// TwinCAT 3 PLC project PannenkoekSysteem
// ProgramVersion: 3.1.4026.20
// CompilerDefines: VISU_USEPROPERTYINFO
// libraries:
//   Tc2_Standard, * (Beckhoff Automation GmbH)
//   Tc2_System, * (Beckhoff Automation GmbH)
//   Tc3_IotBase, * (Beckhoff Automation GmbH)
//   Tc3_Module, * (Beckhoff Automation GmbH)
//   Tc3_Vision, * (Beckhoff Automation GmbH)
// project tree:
//   DUTs/ E_MainState.TcDUT
//   / GlobalTextList.TcGTLO, PlcTask.TcTTO, Visualization Manager.TcVMO (not stored)
//   GVLs/ GVL_Config.TcGVL, GVL_Data.TcGVL, GVL_Inputs.TcGVL, GVL_MQTT.TcGVL, GVL_Outputs.TcGVL
//   POUs/ FB_MQTT.TcPOU, FB_QrVision.TcPOU, F_ParseErrorDisplay.TcPOU, F_ParseStateDisplay.TcPOU, FB_StateMachine.TcPOU, FB_Transportband.TcPOU, MAIN.TcPOU
//   VISUs/ PannenkoekenDashboard.TcVIS
// real-time tasks:
//   TASK PlcTask: cycle T#10ms, priority 20, ADS port 350
//   TASK VnTask ImgAcq (Camera1): cycle T#1ms, priority 5, ADS port 351
//   TASK VnTask ADS (Camera1): cycle T#10ms, priority 6, ADS port 352
// motion (NC):
//   TASK NC-Task 1 SAF: cycle T#2ms, priority 4, ADS port 501
//   TASK NC-Task 1 SVB: cycle T#10ms, priority 8, ADS port 511
//   AXIS Axis 1 (id 1)
//     Dynamic: AccelerationMaximum=200, DecelerationMaximum=200
//     Velo: SlowManual=5, FastManual=20, Maximum=50
//     MotionControl: Range=500, Time=20
//     OtherSettings: AllowMotionCmdToSlave=true
//     encoder EncType=4
//       EncPara: EncMode=1, MaxCount=#x0000ffff
//     drive DrvType=23
//       Analog: VeloReferenz=50, TorqueSetpointScale=10, ScaleFactorActTorque=0.1
//       TimeComp: TaskDelayCycles=1
//     controller CtrType=1
//       CtrPara: PriorControlFactor=1
//         PosDiffControl: Range=20000
//         Observer: BandWidth=20
// I/O:
//   DEVICE Device 2 (EtherCAT), AmsNetId 172.18.237.156.3.1
//     Term 1 (EK1100) [EK1100 EtherCAT Coupler (2A E-Bus)]
//       Term 2 (EL7332) [EL7332 2Ch. DC motor output stage (24V, 1.5A)]
//       Term 3 (EL6001) [EL6001 Interface (RS232)]
//       Box 4 (BK1250)
//   DEVICE Device 1 (RT-Ethernet Adapter)
// variable links:
//   NC-Task 1 SAF/Axes/Axis 1 <-> Device 2 (EtherCAT)/Term 1 (EK1100)/Term 2 (EL7332)
//     Drive/Inputs/In/nState1 @bit 3 <-> DCM Status Channel 1/Status/Error
//     Drive/Inputs/In/nState1 @bit 5 <-> DCM Status Channel 1/Status/Moving negative
//     Drive/Inputs/In/nState1 @bit 4 <-> DCM Status Channel 1/Status/Moving positive
//     Drive/Inputs/In/nState1 @bit 1 <-> DCM Status Channel 1/Status/Ready
//     Drive/Inputs/In/nState1 <-> DCM Status Channel 1/Status/Ready to enable
//     Drive/Inputs/In/nState1 @bit 6 <-> DCM Status Channel 1/Status/Torque reduced
//     Drive/Inputs/In/nState1 @bit 2 <-> DCM Status Channel 1/Status/Warning
//     Drive/Inputs/In/nState2 @bit 3 <-> DCM Status Channel 1/Status/Digital input 1
//     Drive/Inputs/In/nState2 @bit 4 <-> DCM Status Channel 1/Status/Digital input 2
//     Drive/Inputs/In/nState2 @bit 5 <-> DCM Status Channel 1/Status/Sync error
//     Drive/Inputs/In/nState2 @bit 7 <-> DCM Status Channel 1/Status/TxPDO Toggle
//     Drive/Inputs/In/nState4 @bit 1 <-> WcState/InputToggle
//     Drive/Inputs/In/nState4 <-> WcState/WcState
//     Drive/Outputs/Out/nCtrl1 <-> DCM Control Channel 1/Control/Enable
//     Drive/Outputs/Out/nCtrl1 @bit 2 <-> DCM Control Channel 1/Control/Reduce torque
//     Drive/Outputs/Out/nCtrl1 @bit 1 <-> DCM Control Channel 1/Control/Reset
//     Drive/Outputs/Out/nDataOut2[0] <-> DCM Velocity Channel 1/Velocity

CONFIGURATION PannenkoekSysteem
    RESOURCE PLC ON TwinCAT3
        TASK PlcTask(INTERVAL := T#10ms, PRIORITY := 20);
        PROGRAM MAIN WITH PlcTask : MAIN;
    END_RESOURCE
END_CONFIGURATION

// ---- DUTs/E_MainState.TcDUT
{attribute 'qualified_only'}
{attribute 'strict'}
TYPE E_MainState :
(
    INIT,
    IDLE,
    ERROR,
    SEQ_WAIT_START,
    SEQ_FEED_BLOCK,
    SEQ_MOVE_CAMERA,
    SEQ_WAIT_CAMERA,
    SEQ_SCAN_CAMERA,
    SEQ_MOVE_SCALE,
    SEQ_WAIT_SCALE,
    SEQ_MOVE_MIXER,
    SEQ_WAIT_MIXER,
    SEQ_MOVE_INDUCTIVE,
    SEQ_WAIT_INDUCTIVE,
    SEQ_MOVE_DISCARD,
    SEQ_WAIT_DISCARD,
    SEQ_COMPLETE,
    SEQ_ERROR
);
END_TYPE

// ---- GVLs/GVL_Config.TcGVL
{attribute 'qualified_only'}
VAR_GLOBAL
  bAutoSequenceEnable : BOOL := TRUE;      // Master switch for the automated line sequence
  tFeedDuration       : TIME := T#3S;      // Conveyor run time before the robot starts
  tRobotTimeout       : TIME := T#20S;     // Max time to wait for a robot move
  tQrScanDuration     : TIME := T#5S;      // Max time to scan the block at the camera
  tSensorWaitDuration : TIME := T#5S;      // Max time to wait for the inductive sensor

  sPoseCamera    : STRING(32) := 'camera';
  sPoseScale     : STRING(32) := 'scale';
  sPoseMixer     : STRING(32) := 'mixer';
  sPoseInductive : STRING(32) := 'inductive';
  sPoseDiscard   : STRING(32) := 'discard';
END_VAR

// ---- GVLs/GVL_Data.TcGVL
{attribute 'qualified_only'}
VAR_GLOBAL
  bQrEnabled     : BOOL := FALSE;
  bQrCodeFound   : BOOL := FALSE;
  bQrCameraConnected : BOOL := FALSE; // Camera hardware connected
  bQrActive      : BOOL := FALSE;    // Enabled OR camera connected (VISU lamp)
  sQrCodeText    : STRING(255) := '';
  sQrDisplayText : STRING(512) := 'QR scanner OFF';
  hrQrVision     : HRESULT := 0;
END_VAR

// ---- GVLs/GVL_Inputs.TcGVL
{attribute 'qualified_only'}
  VAR_GLOBAL
  END_VAR

// ---- GVLs/GVL_MQTT.TcGVL
{attribute 'qualified_only'}
VAR_GLOBAL
	// MQTT Broker Configuration - HiveMQ Public Broker
	sMqttBroker			: STRING(255) := '192.168.0.198';	// MQTT broker address
	nMqttPort			: UINT := 1883;						// Standard MQTT port
	sMqttClientID		: STRING(255) := 'Twincat_Test'; // Unique client ID
	bEnableMqtt			: BOOL := TRUE;						// Enable/disable MQTT connection
	
	// MQTT Topics - Robot
	sTopicRobotCmd			: STRING(255) := 'pancake/robot/cmd';
	sTopicRobotState		: STRING(255) := 'pancake/robot/state';
	sTopicRobotError		: STRING(255) := 'pancake/robot/error';
	sTopicRobotHeartbeat	: STRING(255) := 'pancake/robot/heartbeat';

	// MQTT Topics - Transportband
	sTopicTransportbandCmd		: STRING(255) := 'pancake/transportband/cmd';
	sTopicTransportbandState	: STRING(255) := 'pancake/transportband/state';
	sTopicTransportbandError	: STRING(255) := 'pancake/transportband/error';

	// MQTT Topics - Mixer
	sTopicMixerCmd				: STRING(255) := 'pancake/mixer/cmd';
	sTopicMixerState			: STRING(255) := 'pancake/mixer/state';
	sTopicMixerError			: STRING(255) := 'pancake/mixer/error';
	
	bVisuStartTransportband : BOOL := FALSE;				// VISU button - Start transportband
	bVisuStopTransportband	: BOOL := FALSE;				// VISU button - Stop transportband
	bVisuStartSequence		: BOOL := FALSE;				// VISU button - Start automated sequence
	bVisuAutoSequenceEnable	: BOOL := TRUE;				// VISU toggle - Automatic line sequence
	
	bVisuStartRobotArm		: BOOL := FALSE;				// Legacy: go-to selected pose
	bVisuStopRobotArm		: BOOL := FALSE;				// Legacy: robot stop
	bVisuRobotTeach			: BOOL := FALSE;				// Teach selected pose
	bVisuRobotGoto				: BOOL := FALSE;				// Go-to selected pose
	bVisuRobotSave				: BOOL := FALSE;				// Save current teach step
	bVisuRobotStop				: BOOL := FALSE;				// Stop/abort robot
	sRobotTargetPose			: STRING(32) := 'camera';	// Target pose for teach/goto

	bVisuForceDisableTeachIndicator : BOOL := FALSE;
	
	// Status variables
	bMqttConnected		: BOOL := FALSE;
	sCurrentState		: STRING(255) := 'IDLE';
	bRobotArmOnline		: BOOL := FALSE;
	bRobotArmRunning		: BOOL := FALSE;
	bRobotArmBusy			: BOOL := FALSE;
	bRobotArmTeachMode		: BOOL := FALSE;
	bRobotArmAlarm			: BOOL := FALSE;
	bRobotArmAckOk			: BOOL := FALSE;
	bRobotArmDone			: BOOL := FALSE;
	sRobotArmDisplay		: STRING(255) := 'Robot Arm OFFLINE';
	sRobotArmAck			: STRING(255) := '';
	sRobotArmLastCommand	: STRING(255) := '';
	sRobotArmLastPose		: STRING(32) := '';
	sRobotHeartbeatRaw		: STRING(255) := '';
	sRobotHeartbeatDisplay	: STRING(255) := '';
	bTransportbandRunning : BOOL := FALSE;
	bTransportbandDone	: BOOL := FALSE;
	sTransportbandDisplay : STRING(255) := 'Transportband OFF';
	bSystemError		: BOOL := FALSE;
	sErrorMessage		: STRING(255) := '';

	// Robot data (READ ONLY via Subscribe)
	{attribute 'TcEncoding':='UTF-8'}
	sRobotCmdRaw		: STRING(255) := '';
	{attribute 'TcEncoding':='UTF-8'}
	sRobotStateRaw		: STRING(255) := '';
	{attribute 'TcEncoding':='UTF-8'}
	sRobotErrorRaw		: STRING(255) := '';
	{attribute 'TcEncoding':='UTF-8'}
	sRobotCmdDisplay	: STRING(255) := '';
	{attribute 'TcEncoding':='UTF-8'}
	sRobotStateDisplay	: STRING(255) := '';
	{attribute 'TcEncoding':='UTF-8'}
	sRobotErrorDisplay	: STRING(255) := '';
	{attribute 'TcEncoding':='UTF-8'}
	sTransportbandCmdRaw : STRING(255) := '';
	{attribute 'TcEncoding':='UTF-8'}
	sMixerCmdRaw		: STRING(255) := '';
	{attribute 'TcEncoding':='UTF-8'}
	sMixerStateRaw		: STRING(255) := '';
	{attribute 'TcEncoding':='UTF-8'}
	sMixerErrorRaw		: STRING(255) := '';
	{attribute 'TcEncoding':='UTF-8'}
	sMixerCmdDisplay	: STRING(255) := '';
	{attribute 'TcEncoding':='UTF-8'}
	sMixerStateDisplay	: STRING(255) := '';
	{attribute 'TcEncoding':='UTF-8'}
	sMixerErrorDisplay	: STRING(255) := '';
	
END_VAR

// ---- GVLs/GVL_Outputs.TcGVL
{attribute 'qualified_only'}
VAR_GLOBAL
END_VAR

// ---- POUs/MAIN.TcPOU
PROGRAM MAIN
VAR
  fbStateMachine    : FB_StateMachine;
  fbTransportband   : FB_Transportband;
  fbMqtt            : FB_MQTT;
  fbQrVision        : FB_QrVision;
  rVisuStartTap     : R_TRIG;
  rVisuStopTap      : R_TRIG;
  rRobotTeachTap    : R_TRIG;
  rRobotGotoTap     : R_TRIG;
  rRobotSaveTap     : R_TRIG;
  rRobotStopTap     : R_TRIG;

  bStartRequest     : BOOL := FALSE;
  bStopRequest      : BOOL := FALSE;
  bStartCmd         : BOOL := FALSE;
  bStopCmd          : BOOL := FALSE;
  bRobotTeachCmd    : BOOL := FALSE;
  bRobotGotoCmd     : BOOL := FALSE;
  bRobotSaveCmd     : BOOL := FALSE;
  bRobotStopCmd     : BOOL := FALSE;
  
  // Transportband - Inductive sensor and DC motor control (EL7332)
  bInductiveSensor  : BOOL := FALSE;   // Inductive sensor input (digital input terminal)
  nMotorOutput      : INT := 0;        // Motor output for DC motor via EL7332 (0-32767 = 0-10V)
END_VAR

// 1) Start/stop requests for the line
rVisuStartTap(CLK := GVL_MQTT.bVisuStartTransportband OR GVL_MQTT.bVisuStartSequence);
rVisuStopTap(CLK := GVL_MQTT.bVisuStopTransportband);

// If the user presses the Start Sequence button, enable AUTO and start immediately
IF rVisuStartTap.Q THEN
  GVL_MQTT.bVisuAutoSequenceEnable := TRUE;
  GVL_Config.bAutoSequenceEnable := TRUE;
END_IF

// Config follows VISU toggle
GVL_Config.bAutoSequenceEnable := GVL_MQTT.bVisuAutoSequenceEnable;

bStartRequest := rVisuStartTap.Q OR fbMqtt.bRemoteStart;
bStopRequest := rVisuStopTap.Q OR fbMqtt.bRemoteStop;

// 2) State machine owns the automation sequence
fbStateMachine(
  bAutoEnable := GVL_Config.bAutoSequenceEnable,
  bStartRequest := bStartRequest,
  bStopRequest := bStopRequest,
  bError := GVL_MQTT.bSystemError,
  bTransportbandDone := fbTransportband.bDone,
  bRobotBusy := fbMqtt.bRobotArmBusy,
  bRobotDone := fbMqtt.bRobotArmDone,
  bQrCodeFound := GVL_Data.bQrCodeFound,
  bInductiveSensor := bInductiveSensor,
  tRobotTimeout := GVL_Config.tRobotTimeout,
  tQrScanDuration := GVL_Config.tQrScanDuration,
  tSensorWaitDuration := GVL_Config.tSensorWaitDuration,
  sPoseCamera := GVL_Config.sPoseCamera,
  sPoseScale := GVL_Config.sPoseScale,
  sPoseMixer := GVL_Config.sPoseMixer,
  sPoseInductive := GVL_Config.sPoseInductive,
  sPoseDiscard := GVL_Config.sPoseDiscard
);

  bStartCmd := fbStateMachine.bStartCmd;
  bStopCmd := fbStateMachine.bStopCmd;
  bRobotGotoCmd := fbStateMachine.bRobotGotoCmd;
  bRobotStopCmd := fbStateMachine.bRobotStopCmd;
  bRobotTeachCmd := FALSE;
  bRobotSaveCmd := FALSE;

  IF NOT GVL_Config.bAutoSequenceEnable THEN
    // Manual robot controls remain available when automation is disabled
    rRobotTeachTap(CLK := GVL_MQTT.bVisuRobotTeach);
    rRobotGotoTap(CLK := GVL_MQTT.bVisuRobotGoto OR GVL_MQTT.bVisuStartRobotArm);
    rRobotSaveTap(CLK := GVL_MQTT.bVisuRobotSave);
    rRobotStopTap(CLK := GVL_MQTT.bVisuRobotStop OR GVL_MQTT.bVisuStopRobotArm);

    IF rRobotStopTap.Q THEN
      bRobotStopCmd := TRUE;
    ELSIF rRobotSaveTap.Q THEN
      bRobotSaveCmd := TRUE;
    ELSIF rRobotTeachTap.Q THEN
      bRobotTeachCmd := TRUE;
    ELSIF rRobotGotoTap.Q THEN
      bRobotGotoCmd := TRUE;
    END_IF

    bStartCmd := bStartRequest;
    bStopCmd := bStopRequest;
  END_IF

  // Clear VISU request flags so each button click becomes a fresh rising edge
  GVL_MQTT.bVisuRobotTeach := FALSE;
  GVL_MQTT.bVisuRobotGoto  := FALSE;
  GVL_MQTT.bVisuRobotSave  := FALSE;
  GVL_MQTT.bVisuRobotStop  := FALSE;
  GVL_MQTT.bVisuStartRobotArm := FALSE;
  GVL_MQTT.bVisuStopRobotArm  := FALSE;
  GVL_MQTT.bVisuStartSequence := FALSE;

  // Update robot arm status display from MQTT feedback
  GVL_MQTT.bRobotArmOnline := fbMqtt.bRobotArmOnline;
  GVL_MQTT.bRobotArmRunning := fbMqtt.bRobotArmRunning;
  GVL_MQTT.bRobotArmBusy := fbMqtt.bRobotArmBusy;
  GVL_MQTT.bRobotArmTeachMode := fbMqtt.bRobotArmTeachMode;
  GVL_MQTT.bRobotArmAlarm := fbMqtt.bRobotArmAlarm;
  GVL_MQTT.bRobotArmDone := fbMqtt.bRobotArmDone;
  GVL_MQTT.bRobotArmAckOk := fbMqtt.bRobotArmAckOk;

  IF NOT GVL_MQTT.bRobotArmOnline THEN
    GVL_MQTT.sRobotArmDisplay := 'Robot Arm OFFLINE';
  ELSIF GVL_MQTT.bRobotArmAlarm THEN
    GVL_MQTT.sRobotArmDisplay := 'Robot Arm ALARM';
  ELSIF GVL_MQTT.bRobotArmTeachMode THEN
    GVL_MQTT.sRobotArmDisplay := 'Robot Arm TEACH';
  ELSIF GVL_MQTT.bRobotArmBusy THEN
    GVL_MQTT.sRobotArmDisplay := 'Robot Arm BUSY';
  ELSIF GVL_MQTT.bRobotArmDone THEN
    GVL_MQTT.sRobotArmDisplay := 'Robot Arm READY';
  ELSE
    GVL_MQTT.sRobotArmDisplay := 'Robot Arm READY';
  END_IF

  GVL_MQTT.sCurrentState := TO_STRING(fbStateMachine.eStateOut);

  // 3) Transportband
  fbTransportband(
    bStart := bStartCmd,
    bStop := bStopCmd,
    tDuration := GVL_Config.tFeedDuration
  );

  GVL_MQTT.bTransportbandRunning := fbTransportband.bRunning;
  GVL_MQTT.bTransportbandDone := fbTransportband.bDone;
  nMotorOutput := fbTransportband.nMotorControl;

  IF fbTransportband.bRunning THEN
    GVL_MQTT.sTransportbandDisplay := 'Transportband ON';
  ELSIF fbTransportband.bDone THEN
    GVL_MQTT.sTransportbandDisplay := 'Transportband READY';
  ELSE
    GVL_MQTT.sTransportbandDisplay := 'Transportband OFF';
  END_IF

  // 4) MQTT in separate function block
  fbMqtt(
    bTransportbandRunning := GVL_MQTT.bTransportbandRunning,
    bTransportbandDone := GVL_MQTT.bTransportbandDone,
    bRobotTeachCmd := bRobotTeachCmd,
    bRobotGotoCmd := bRobotGotoCmd,
    bRobotSaveCmd := bRobotSaveCmd,
    bRobotStopCmd := bRobotStopCmd,
    sRobotTargetPose := GVL_MQTT.sRobotTargetPose,
    bSystemError := GVL_MQTT.bSystemError,
    sErrorMessage := GVL_MQTT.sErrorMessage
  );

  // 5) QR vision
  fbQrVision(
    bEnable := GVL_Data.bQrEnabled OR fbStateMachine.bQrAutoEnable
  );

  GVL_Data.bQrCodeFound := fbQrVision.bCodeFound;
  GVL_Data.sQrCodeText := fbQrVision.sCodeAsString;
  GVL_Data.sQrDisplayText := fbQrVision.sDisplayText;
  GVL_Data.hrQrVision := fbQrVision.hrLast;

  // Expose camera connected state and combined active flag for VISU
  GVL_Data.bQrCameraConnected := fbQrVision.bCameraConnected;
  GVL_Data.bQrActive := GVL_Data.bQrEnabled OR fbQrVision.bCameraConnected;

END_PROGRAM

// ---- POUs/FB_StateMachine.TcPOU
FUNCTION_BLOCK FB_StateMachine

VAR_INPUT
    bAutoEnable         : BOOL := TRUE;
    bStartRequest       : BOOL;
    bStopRequest        : BOOL;
    bError              : BOOL;
    bTransportbandDone  : BOOL;
    bRobotBusy          : BOOL;
    bRobotDone          : BOOL;
    bQrCodeFound        : BOOL;
    bInductiveSensor    : BOOL;
    tRobotTimeout       : TIME;
    tQrScanDuration     : TIME;
    tSensorWaitDuration : TIME;
    sPoseCamera         : STRING(32);
    sPoseScale          : STRING(32);
    sPoseMixer          : STRING(32);
    sPoseInductive      : STRING(32);
    sPoseDiscard        : STRING(32);
END_VAR

VAR_OUTPUT
    eStateOut         : E_MainState; // Current state visible outside
    bStartCmd         : BOOL;
    bStopCmd          : BOOL;
    bRobotGotoCmd     : BOOL;
    bRobotStopCmd     : BOOL;
    bQrAutoEnable     : BOOL;
    sRobotTargetPose  : STRING(32);
END_VAR

VAR
	eState : E_MainState := E_MainState.INIT;
	bRobotBusySeen : BOOL := FALSE;
	tRobotTimeoutFb : TON;
	tQrScanTimerFb : TON;
	tSensorWaitTimerFb : TON;
END_VAR

// Default outputs
bStartCmd := FALSE;
bStopCmd := FALSE;
bRobotGotoCmd := FALSE;
bRobotStopCmd := FALSE;
bQrAutoEnable := FALSE;
sRobotTargetPose := '';

// Reset timers unless the active state enables them below
tRobotTimeoutFb(IN := FALSE, PT := tRobotTimeout);
tQrScanTimerFb(IN := FALSE, PT := tQrScanDuration);
tSensorWaitTimerFb(IN := FALSE, PT := tSensorWaitDuration);

CASE eState OF
  E_MainState.INIT:
    eState := E_MainState.IDLE;

  E_MainState.IDLE:
    IF bError THEN
      eState := E_MainState.ERROR;
    ELSIF bAutoEnable AND bStartRequest THEN
      eState := E_MainState.SEQ_FEED_BLOCK;
      bRobotBusySeen := FALSE;
    END_IF

  E_MainState.SEQ_FEED_BLOCK:
    bStartCmd := TRUE;
    IF bStopRequest OR bError THEN
      eState := E_MainState.SEQ_ERROR;
    ELSIF bTransportbandDone THEN
      eState := E_MainState.SEQ_MOVE_CAMERA;
    END_IF

  E_MainState.SEQ_MOVE_CAMERA:
    bRobotGotoCmd := TRUE;
    sRobotTargetPose := sPoseCamera;
    eState := E_MainState.SEQ_WAIT_CAMERA;

  E_MainState.SEQ_WAIT_CAMERA:
    tRobotTimeoutFb(IN := TRUE, PT := tRobotTimeout);
    IF bError OR bStopRequest THEN
      eState := E_MainState.SEQ_ERROR;
    ELSE
      IF bRobotBusy THEN
        bRobotBusySeen := TRUE;
      END_IF

      IF bRobotBusySeen AND bRobotDone AND NOT bRobotBusy THEN
        bRobotBusySeen := FALSE;
        eState := E_MainState.SEQ_SCAN_CAMERA;
      ELSIF tRobotTimeoutFb.Q THEN
        eState := E_MainState.SEQ_ERROR;
      END_IF
    END_IF

  E_MainState.SEQ_SCAN_CAMERA:
    bQrAutoEnable := TRUE;
    tQrScanTimerFb(IN := TRUE, PT := tQrScanDuration);
    IF bQrCodeFound OR tQrScanTimerFb.Q THEN
      eState := E_MainState.SEQ_MOVE_SCALE;
    END_IF

  E_MainState.SEQ_MOVE_SCALE:
    bRobotGotoCmd := TRUE;
    sRobotTargetPose := sPoseScale;
    eState := E_MainState.SEQ_WAIT_SCALE;

  E_MainState.SEQ_WAIT_SCALE:
    tRobotTimeoutFb(IN := TRUE, PT := tRobotTimeout);
    IF bError OR bStopRequest THEN
      eState := E_MainState.SEQ_ERROR;
    ELSE
      IF bRobotBusy THEN
        bRobotBusySeen := TRUE;
      END_IF

      IF bRobotBusySeen AND bRobotDone AND NOT bRobotBusy THEN
        bRobotBusySeen := FALSE;
        eState := E_MainState.SEQ_MOVE_MIXER;
      ELSIF tRobotTimeoutFb.Q THEN
        eState := E_MainState.SEQ_ERROR;
      END_IF
    END_IF

  E_MainState.SEQ_MOVE_MIXER:
    bRobotGotoCmd := TRUE;
    sRobotTargetPose := sPoseMixer;
    eState := E_MainState.SEQ_WAIT_MIXER;

  E_MainState.SEQ_WAIT_MIXER:
    tRobotTimeoutFb(IN := TRUE, PT := tRobotTimeout);
    IF bError OR bStopRequest THEN
      eState := E_MainState.SEQ_ERROR;
    ELSE
      IF bRobotBusy THEN
        bRobotBusySeen := TRUE;
      END_IF

      IF bRobotBusySeen AND bRobotDone AND NOT bRobotBusy THEN
        bRobotBusySeen := FALSE;
        eState := E_MainState.SEQ_MOVE_INDUCTIVE;
      ELSIF tRobotTimeoutFb.Q THEN
        eState := E_MainState.SEQ_ERROR;
      END_IF
    END_IF

  E_MainState.SEQ_MOVE_INDUCTIVE:
    bRobotGotoCmd := TRUE;
    sRobotTargetPose := sPoseInductive;
    eState := E_MainState.SEQ_WAIT_INDUCTIVE;

  E_MainState.SEQ_WAIT_INDUCTIVE:
    tRobotTimeoutFb(IN := TRUE, PT := tRobotTimeout);
    IF bError OR bStopRequest THEN
      eState := E_MainState.SEQ_ERROR;
    ELSE
      IF bRobotBusy THEN
        bRobotBusySeen := TRUE;
      END_IF

      IF bRobotBusySeen AND bRobotDone AND NOT bRobotBusy THEN
        bRobotBusySeen := FALSE;
        IF bInductiveSensor THEN
          eState := E_MainState.SEQ_MOVE_DISCARD;
        ELSE
          tSensorWaitTimerFb(IN := TRUE, PT := tSensorWaitDuration);
          IF tSensorWaitTimerFb.Q THEN
            eState := E_MainState.SEQ_MOVE_DISCARD;
          END_IF
        END_IF
      ELSIF tRobotTimeoutFb.Q THEN
        eState := E_MainState.SEQ_ERROR;
      END_IF
    END_IF

  E_MainState.SEQ_MOVE_DISCARD:
    bRobotGotoCmd := TRUE;
    sRobotTargetPose := sPoseDiscard;
    eState := E_MainState.SEQ_WAIT_DISCARD;

  E_MainState.SEQ_WAIT_DISCARD:
    tRobotTimeoutFb(IN := TRUE, PT := tRobotTimeout);
    IF bError OR bStopRequest THEN
      eState := E_MainState.SEQ_ERROR;
    ELSE
      IF bRobotBusy THEN
        bRobotBusySeen := TRUE;
      END_IF

      IF bRobotBusySeen AND bRobotDone AND NOT bRobotBusy THEN
        bRobotBusySeen := FALSE;
        eState := E_MainState.SEQ_COMPLETE;
      ELSIF tRobotTimeoutFb.Q THEN
        eState := E_MainState.SEQ_ERROR;
      END_IF
    END_IF

  E_MainState.SEQ_COMPLETE:
    eState := E_MainState.IDLE;

  E_MainState.ERROR:
    bStopCmd := TRUE;
    bRobotStopCmd := TRUE;
    IF bStopRequest THEN
      eState := E_MainState.IDLE;
    END_IF

  E_MainState.SEQ_ERROR:
    bStopCmd := TRUE;
    bRobotStopCmd := TRUE;
    IF bStopRequest THEN
      eState := E_MainState.IDLE;
    END_IF
END_CASE

eStateOut := eState;

END_FUNCTION_BLOCK

// ---- POUs/FB_Transportband.TcPOU
FUNCTION_BLOCK FB_Transportband

VAR_INPUT
    bStart   : BOOL;   // Signal from state machine - start motor
    bStop    : BOOL;   // Stop / emergency stop
    tDuration : TIME;  // Motor run duration
END_VAR

VAR_OUTPUT
    bRunning : BOOL;   // Transportband running
    bDone    : BOOL;   // Transportband cycle complete
    nMotorControl : INT;  // Output for EL7332 DC motor (0-32767 = 0-10V)
END_VAR

VAR
  tRun : TON;       // Timer for motor duration
  rStartTrig : R_TRIG;
  bCycleActive : BOOL := FALSE;
END_VAR

rStartTrig(CLK := bStart);

IF bStop THEN
  // Emergency stop - shut down everything
  bCycleActive := FALSE;
  bRunning := FALSE;
  bDone := FALSE;
  nMotorControl := 0;
  tRun(IN := FALSE);
ELSE
  // New cycle on rising edge of start
  IF rStartTrig.Q THEN
    bDone := FALSE;
    bCycleActive := TRUE;
    nMotorControl := 32767;  // Motor at max speed (10V on EL7332)
  END_IF

  IF bCycleActive THEN
    bRunning := TRUE;
    tRun(IN := TRUE, PT := tDuration);

    // Cycle completes when timer expires
    IF tRun.Q THEN
      bCycleActive := FALSE;
      bRunning := FALSE;
      bDone := TRUE;
      nMotorControl := 0;  // Motor stopped
      tRun(IN := FALSE);
    END_IF
  ELSE
    bRunning := FALSE;
    nMotorControl := 0;  // Motor stopped when no cycle active
    tRun(IN := FALSE);
  END_IF
END_IF

END_FUNCTION_BLOCK

// ---- POUs/FB_MQTT.TcPOU
FUNCTION_BLOCK FB_MQTT
VAR_INPUT
	bTransportbandRunning	: BOOL;
	bTransportbandDone		: BOOL;
	bRobotTeachCmd			: BOOL;
	bRobotGotoCmd			: BOOL;
	bRobotSaveCmd			: BOOL;
	bRobotStopCmd			: BOOL;
	{attribute 'TcEncoding':='UTF-8'}
	sRobotTargetPose		: STRING(32);
	bSystemError			: BOOL;
	{attribute 'TcEncoding':='UTF-8'}
	sErrorMessage			: STRING(255);
END_VAR

VAR_OUTPUT
	bRemoteStart			: BOOL;
	bRemoteStop			: BOOL;
	bRemoteRobotTeach		: BOOL;
	bRemoteRobotGoto		: BOOL;
	bRemoteRobotSave		: BOOL;
	bRemoteRobotStop		: BOOL;
	bRobotArmRunning		: BOOL;
	bRobotArmDone			: BOOL;
	bRobotArmOnline			: BOOL;
	bRobotArmBusy			: BOOL;
	bRobotArmTeachMode		: BOOL;
	bRobotArmAlarm			: BOOL;
	bRobotArmAckOk			: BOOL;
END_VAR

VAR
	fbMqttClient			: FB_IotMqttClient;
	fbMessageQueue			: FB_IotMqttMessageQueue;
	fbMessage				: FB_IotMqttMessage;

	bMqttConfigured			: BOOL := FALSE;
	bSubscribedRobotCmd		: BOOL := FALSE;
	bSubscribedRobotState	: BOOL := FALSE;
	bSubscribedRobotError	: BOOL := FALSE;
	bSubscribedRobotHeartbeat	: BOOL := FALSE;
	bSubscribedTransportState	: BOOL := FALSE;
	bSubscribedMixerCmd		: BOOL := FALSE;
	bSubscribedMixerState	: BOOL := FALSE;
	bSubscribedMixerError	: BOOL := FALSE;
	bSubscribedTransportCmd	: BOOL := FALSE;

	{attribute 'TcEncoding':='UTF-8'}
	sPayloadRcv			: STRING(255);
	{attribute 'TcEncoding':='UTF-8'}
	sPayloadPub			: STRING(255);
	{attribute 'TcEncoding':='UTF-8'}
	sTransportState			: STRING(64);
	{attribute 'TcEncoding':='UTF-8'}
	sRobotState				: STRING(64);
	{attribute 'TcEncoding':='UTF-8'}
	sRobotCommandPayload	: STRING(255);
	{attribute 'TcEncoding':='UTF-8'}
	sLastStatePayload		: STRING(255);
	{attribute 'TcEncoding':='UTF-8'}
	sLastErrorPayload		: STRING(255);
	{attribute 'TcEncoding':='UTF-8'}
	sLastRobotStatePayload	: STRING(255);
	bStatePublished			: BOOL := FALSE;
	bErrorPublished			: BOOL := FALSE;
	bRobotStatePublished	: BOOL := FALSE;
	bRobotHeartbeatPulse	: BOOL := FALSE;
	bRobotStateReceived		: BOOL := FALSE;
	bRobotErrorActive		: BOOL := FALSE;
	fbRobotHeartbeatWatchdog	: TON;
END_VAR

IF NOT bMqttConfigured THEN
	bMqttConfigured := TRUE;
	fbMqttClient.sHostName := GVL_MQTT.sMqttBroker;
	fbMqttClient.nHostPort := GVL_MQTT.nMqttPort;
	fbMqttClient.sClientId := GVL_MQTT.sMqttClientID;
	fbMqttClient.ipMessageQueue := fbMessageQueue;
END_IF

fbMqttClient.Execute(bConnect := GVL_MQTT.bEnableMqtt);
GVL_MQTT.bMqttConnected := fbMqttClient.bConnected;

IF fbMqttClient.bConnected THEN
	IF NOT bSubscribedRobotCmd THEN
		bSubscribedRobotCmd := fbMqttClient.Subscribe(
			sTopic := GVL_MQTT.sTopicRobotCmd,
			eQoS := TcIotMqttQos.AtMostOnceDelivery
		);
	END_IF

	IF NOT bSubscribedRobotState THEN
		bSubscribedRobotState := fbMqttClient.Subscribe(
			sTopic := GVL_MQTT.sTopicRobotState,
			eQoS := TcIotMqttQos.AtMostOnceDelivery
		);
	END_IF

	IF NOT bSubscribedRobotError THEN
		bSubscribedRobotError := fbMqttClient.Subscribe(
			sTopic := GVL_MQTT.sTopicRobotError,
			eQoS := TcIotMqttQos.AtMostOnceDelivery
		);
	END_IF

	IF NOT bSubscribedRobotHeartbeat THEN
		bSubscribedRobotHeartbeat := fbMqttClient.Subscribe(
			sTopic := GVL_MQTT.sTopicRobotHeartbeat,
			eQoS := TcIotMqttQos.AtMostOnceDelivery
		);
	END_IF

	IF NOT bSubscribedTransportState THEN
		bSubscribedTransportState := fbMqttClient.Subscribe(
			sTopic := GVL_MQTT.sTopicTransportbandState,
			eQoS := TcIotMqttQos.AtMostOnceDelivery
		);
	END_IF

	IF NOT bSubscribedMixerCmd THEN
		bSubscribedMixerCmd := fbMqttClient.Subscribe(
			sTopic := GVL_MQTT.sTopicMixerCmd,
			eQoS := TcIotMqttQos.AtMostOnceDelivery
		);
	END_IF

	IF NOT bSubscribedMixerState THEN
		bSubscribedMixerState := fbMqttClient.Subscribe(
			sTopic := GVL_MQTT.sTopicMixerState,
			eQoS := TcIotMqttQos.AtMostOnceDelivery
		);
	END_IF

	IF NOT bSubscribedMixerError THEN
		bSubscribedMixerError := fbMqttClient.Subscribe(
			sTopic := GVL_MQTT.sTopicMixerError,
			eQoS := TcIotMqttQos.AtMostOnceDelivery
		);
	END_IF

	IF NOT bSubscribedTransportCmd THEN
		bSubscribedTransportCmd := fbMqttClient.Subscribe(
			sTopic := GVL_MQTT.sTopicTransportbandCmd,
			eQoS := TcIotMqttQos.AtMostOnceDelivery
		);
	END_IF

	// Robot arm command publishing from PLC
	IF bRobotTeachCmd THEN
		sRobotCommandPayload := '{"cmd":"teach","pose":"';
		sRobotCommandPayload := CONCAT(sRobotCommandPayload, sRobotTargetPose);
		sRobotCommandPayload := CONCAT(sRobotCommandPayload, '"}');
		fbMqttClient.Publish(
			sTopic := GVL_MQTT.sTopicRobotCmd,
			pPayload := ADR(sRobotCommandPayload),
			nPayloadSize := TO_UDINT(LEN(sRobotCommandPayload) + 1),
			eQoS := TcIotMqttQos.AtLeastOnceDelivery,
			bRetain := FALSE,
			bQueue := FALSE
		);
		GVL_MQTT.sRobotArmLastCommand := 'teach';
		GVL_MQTT.sRobotArmLastPose := sRobotTargetPose;
		GVL_MQTT.sRobotArmAck := CONCAT('Teach sent: ', sRobotTargetPose);
		GVL_MQTT.bRobotArmAckOk := TRUE;
		bRobotArmBusy := TRUE;
		bRobotArmTeachMode := TRUE;
		bRobotArmRunning := TRUE;
		bRobotArmDone := FALSE;
		bRobotArmAlarm := FALSE;
	END_IF

	IF bRobotGotoCmd THEN
		sRobotCommandPayload := '{"cmd":"goto","pose":"';
		sRobotCommandPayload := CONCAT(sRobotCommandPayload, sRobotTargetPose);
		sRobotCommandPayload := CONCAT(sRobotCommandPayload, '"}');
		fbMqttClient.Publish(
			sTopic := GVL_MQTT.sTopicRobotCmd,
			pPayload := ADR(sRobotCommandPayload),
			nPayloadSize := TO_UDINT(LEN(sRobotCommandPayload) + 1),
			eQoS := TcIotMqttQos.AtLeastOnceDelivery,
			bRetain := FALSE,
			bQueue := FALSE
		);
		GVL_MQTT.sRobotArmLastCommand := 'goto';
		GVL_MQTT.sRobotArmLastPose := sRobotTargetPose;
		GVL_MQTT.sRobotArmAck := CONCAT('Goto sent: ', sRobotTargetPose);
		GVL_MQTT.bRobotArmAckOk := TRUE;
		bRobotArmBusy := TRUE;
		bRobotArmTeachMode := FALSE;
		bRobotArmRunning := TRUE;
		bRobotArmDone := FALSE;
		bRobotArmAlarm := FALSE;
	END_IF

	IF bRobotSaveCmd THEN
		sRobotCommandPayload := '{"cmd":"save"}';
		fbMqttClient.Publish(
			sTopic := GVL_MQTT.sTopicRobotCmd,
			pPayload := ADR(sRobotCommandPayload),
			nPayloadSize := TO_UDINT(LEN(sRobotCommandPayload) + 1),
			eQoS := TcIotMqttQos.AtLeastOnceDelivery,
			bRetain := FALSE,
			bQueue := FALSE
		);
		GVL_MQTT.sRobotArmLastCommand := 'save';
		GVL_MQTT.sRobotArmAck := 'Save sent';
		GVL_MQTT.bRobotArmAckOk := TRUE;
		bRobotArmBusy := TRUE;
		bRobotArmRunning := TRUE;
		bRobotArmDone := FALSE;
		bRobotArmAlarm := FALSE;
	END_IF

	IF bRobotStopCmd THEN
		sRobotCommandPayload := '{"cmd":"stop"}';
		fbMqttClient.Publish(
			sTopic := GVL_MQTT.sTopicRobotCmd,
			pPayload := ADR(sRobotCommandPayload),
			nPayloadSize := TO_UDINT(LEN(sRobotCommandPayload) + 1),
			eQoS := TcIotMqttQos.AtLeastOnceDelivery,
			bRetain := FALSE,
			bQueue := FALSE
		);
		GVL_MQTT.sRobotArmLastCommand := 'stop';
		GVL_MQTT.sRobotArmAck := 'Stop sent';
		GVL_MQTT.bRobotArmAckOk := TRUE;
		bRobotArmBusy := FALSE;
		bRobotArmTeachMode := FALSE;
		bRobotArmRunning := FALSE;
		bRobotArmDone := FALSE;
	END_IF

	IF bSystemError THEN
		sTransportState := 'error';
	ELSIF bTransportbandRunning THEN
		sTransportState := 'running';
	ELSIF bTransportbandDone THEN
		sTransportState := 'done';
	ELSE
		sTransportState := 'idle';
	END_IF

	sPayloadPub := CONCAT('{"state":"', sTransportState);
	sPayloadPub := CONCAT(sPayloadPub, '"}');

	IF (NOT bStatePublished) OR (sPayloadPub <> sLastStatePayload) THEN
		fbMqttClient.Publish(
			sTopic := GVL_MQTT.sTopicTransportbandState,
			pPayload := ADR(sPayloadPub),
			nPayloadSize := TO_UDINT(LEN(sPayloadPub) + 1),
			eQoS := TcIotMqttQos.AtMostOnceDelivery,
			bRetain := FALSE,
			bQueue := FALSE
		);

		sLastStatePayload := sPayloadPub;
		bStatePublished := TRUE;
	END_IF

	IF bSystemError THEN
		sPayloadPub := CONCAT('{"state":"error","error":true,"message":"', sErrorMessage);
		sPayloadPub := CONCAT(sPayloadPub, '"}');
	ELSE
		sPayloadPub := '{"state":"ok","error":false,"message":""}';
	END_IF

	IF (NOT bErrorPublished) OR (sPayloadPub <> sLastErrorPayload) THEN
		fbMqttClient.Publish(
			sTopic := GVL_MQTT.sTopicTransportbandError,
			pPayload := ADR(sPayloadPub),
			nPayloadSize := TO_UDINT(LEN(sPayloadPub) + 1),
			eQoS := TcIotMqttQos.AtMostOnceDelivery,
			bRetain := FALSE,
			bQueue := FALSE
		);

		sLastErrorPayload := sPayloadPub;
		bErrorPublished := TRUE;
	END_IF

	// Robot arm status is built only from received state/error/heartbeat messages.
	// The PLC only publishes commands here, not the robot-state topic.
ELSE
	bSubscribedRobotCmd := FALSE;
	bSubscribedRobotState := FALSE;
	bSubscribedRobotError := FALSE;
	bSubscribedRobotHeartbeat := FALSE;
	bSubscribedTransportState := FALSE;
	bSubscribedMixerCmd := FALSE;
	bSubscribedMixerState := FALSE;
	bSubscribedMixerError := FALSE;
	bSubscribedTransportCmd := FALSE;
	bStatePublished := FALSE;
	bErrorPublished := FALSE;
	bRobotStatePublished := FALSE;
	bRobotArmRunning := FALSE;
	bRobotArmDone := FALSE;
	bRobotArmOnline := FALSE;
	bRobotArmBusy := FALSE;
	bRobotArmTeachMode := FALSE;
	bRobotArmAlarm := FALSE;
	bRobotArmAckOk := FALSE;
	sLastStatePayload := '';
	sLastErrorPayload := '';
	sLastRobotStatePayload := '';
END_IF

// Remote commando's als puls per PLC-cyclus
bRemoteStart := FALSE;
bRemoteStop := FALSE;
bRemoteRobotTeach := FALSE;
bRemoteRobotGoto := FALSE;
bRemoteRobotSave := FALSE;
bRemoteRobotStop := FALSE;

IF fbMessageQueue.nQueuedMessages > 0 THEN
	IF fbMessageQueue.Dequeue(fbMessage := fbMessage) THEN
		fbMessage.GetPayload(
			pPayload := ADR(sPayloadRcv),
			nPayloadSize := SIZEOF(sPayloadRcv),
			bSetNullTermination := FALSE
		);

		IF fbMessage.CompareTopic(sTopic := GVL_MQTT.sTopicRobotCmd) THEN
			GVL_MQTT.sRobotCmdRaw := sPayloadRcv;
			GVL_MQTT.sRobotCmdDisplay := sPayloadRcv;

			IF (FIND(sPayloadRcv, '"cmd":"teach"') > 0) OR (FIND(sPayloadRcv, '"cmd": "teach"') > 0) THEN
				bRemoteRobotTeach := TRUE;
			ELSIF (FIND(sPayloadRcv, '"cmd":"goto"') > 0) OR (FIND(sPayloadRcv, '"cmd": "goto"') > 0) THEN
				bRemoteRobotGoto := TRUE;
			ELSIF (FIND(sPayloadRcv, '"cmd":"save"') > 0) OR (FIND(sPayloadRcv, '"cmd": "save"') > 0) THEN
				bRemoteRobotSave := TRUE;
			ELSIF (FIND(sPayloadRcv, '"cmd":"stop"') > 0) OR (FIND(sPayloadRcv, '"cmd": "stop"') > 0) THEN
				bRemoteRobotStop := TRUE;
			END_IF
		ELSIF fbMessage.CompareTopic(sTopic := GVL_MQTT.sTopicRobotState) THEN
			GVL_MQTT.sRobotStateRaw := sPayloadRcv;
			GVL_MQTT.sRobotStateDisplay := F_ParseStateDisplay(sPayload := sPayloadRcv);
			bRobotStateReceived := TRUE;
			GVL_MQTT.bRobotArmAckOk := TRUE;
			GVL_MQTT.sRobotArmAck := GVL_MQTT.sRobotStateDisplay;

			// Robot sends: teach_<pose>, teach_pose_changed, teach_<pose>_saved_motor*, teach_<pose>_complete, at_<pose>, idle
			IF (FIND(sPayloadRcv, '"state":"teach_') > 0) THEN
				// All teach states → busy in teach mode
				bRobotArmBusy := TRUE;
				bRobotArmTeachMode := TRUE;
				IF (FIND(sPayloadRcv, '"state":"teach_') > 0) AND (FIND(sPayloadRcv, '_complete"') > 0) THEN
					// teach_<pose>_complete → teach done
					bRobotArmDone := TRUE;
					bRobotArmBusy := FALSE;
					bRobotArmRunning := FALSE;
				ELSE
					// teach_<pose>, teach_pose_changed, teach_<pose>_saved_motor* → still teaching
					bRobotArmDone := FALSE;
					bRobotArmRunning := TRUE;
				END_IF
			ELSIF (FIND(sPayloadRcv, '"state":"at_') > 0) THEN
				// at_<pose> → robot reached pose, done
				bRobotArmBusy := FALSE;
				bRobotArmDone := TRUE;
				bRobotArmTeachMode := FALSE;
				bRobotArmRunning := FALSE;
			ELSIF (FIND(sPayloadRcv, '"state":"running"') > 0) THEN
				// running → robot executing action
				bRobotArmBusy := TRUE;
				bRobotArmDone := FALSE;
				bRobotArmTeachMode := FALSE;
				bRobotArmRunning := TRUE;
			ELSIF (FIND(sPayloadRcv, '"state":"done"') > 0) THEN
				// done → action finished
				bRobotArmBusy := FALSE;
				bRobotArmDone := TRUE;
				bRobotArmTeachMode := FALSE;
				bRobotArmRunning := FALSE;
			ELSIF (FIND(sPayloadRcv, '"state":"idle"') > 0) THEN
				// idle → robot at rest
				bRobotArmBusy := FALSE;
				bRobotArmDone := TRUE;
				bRobotArmTeachMode := FALSE;
				bRobotArmRunning := FALSE;
			ELSE
				// Unknown state → stay in previous state to avoid false negatives
				bRobotArmDone := FALSE;
				bRobotArmRunning := FALSE;
			END_IF
		ELSIF fbMessage.CompareTopic(sTopic := GVL_MQTT.sTopicRobotError) THEN
			GVL_MQTT.sRobotErrorRaw := sPayloadRcv;
			GVL_MQTT.sRobotErrorDisplay := F_ParseErrorDisplay(sPayload := sPayloadRcv);
			
			// Robot sends: {"state":"error","error":true,"message":"..."} or {"state":"ok","error":false,"message":""}
			IF (FIND(sPayloadRcv, '"error":true') > 0) THEN
				// Real error
				bRobotErrorActive := TRUE;
				bRobotArmAlarm := TRUE;
				GVL_MQTT.bRobotArmAckOk := FALSE;
				GVL_MQTT.sRobotArmAck := GVL_MQTT.sRobotErrorDisplay;
			ELSE
				// Ok response
				bRobotErrorActive := FALSE;
				bRobotArmAlarm := FALSE;
				GVL_MQTT.bRobotArmAckOk := TRUE;
				GVL_MQTT.sRobotArmAck := 'Robot Error OK';
			END_IF
			bRobotArmRunning := FALSE;
			bRobotArmBusy := FALSE;
		ELSIF fbMessage.CompareTopic(sTopic := GVL_MQTT.sTopicRobotHeartbeat) THEN
			GVL_MQTT.sRobotHeartbeatRaw := sPayloadRcv;
			GVL_MQTT.sRobotHeartbeatDisplay := 'Robot Heartbeat OK';
			bRobotHeartbeatPulse := TRUE;
			GVL_MQTT.bRobotArmOnline := TRUE;
			GVL_MQTT.bRobotArmAckOk := TRUE;
		ELSIF fbMessage.CompareTopic(sTopic := GVL_MQTT.sTopicMixerCmd) THEN
			GVL_MQTT.sMixerCmdRaw := sPayloadRcv;
			GVL_MQTT.sMixerCmdDisplay := sPayloadRcv;
		ELSIF fbMessage.CompareTopic(sTopic := GVL_MQTT.sTopicMixerState) THEN
			GVL_MQTT.sMixerStateRaw := sPayloadRcv;
			GVL_MQTT.sMixerStateDisplay := F_ParseStateDisplay(sPayload := sPayloadRcv);
		ELSIF fbMessage.CompareTopic(sTopic := GVL_MQTT.sTopicMixerError) THEN
			GVL_MQTT.sMixerErrorRaw := sPayloadRcv;
			GVL_MQTT.sMixerErrorDisplay := F_ParseErrorDisplay(sPayload := sPayloadRcv);
		ELSIF fbMessage.CompareTopic(sTopic := GVL_MQTT.sTopicTransportbandCmd) THEN
			GVL_MQTT.sTransportbandCmdRaw := sPayloadRcv;

			IF (sPayloadRcv = '{"cmd":"stop"}') OR (sPayloadRcv = '{"cmd":"STOP"}') OR (sPayloadRcv = 'stop') OR (sPayloadRcv = 'STOP') THEN
				bRemoteStart := FALSE;
				bRemoteStop := TRUE;
			ELSIF (sPayloadRcv = '{"cmd":"start"}') OR (sPayloadRcv = '{"cmd":"START"}') OR (sPayloadRcv = 'start') OR (sPayloadRcv = 'START') THEN
				bRemoteStart := TRUE;
				bRemoteStop := FALSE;
			END_IF
		END_IF
	END_IF
END_IF

fbRobotHeartbeatWatchdog(IN := NOT bRobotHeartbeatPulse, PT := T#12S);
IF fbRobotHeartbeatWatchdog.Q THEN
	GVL_MQTT.bRobotArmOnline := FALSE;
	GVL_MQTT.sRobotHeartbeatDisplay := 'Robot Heartbeat TIMEOUT';
ELSE
	GVL_MQTT.bRobotArmOnline := FALSE;
END_IF
bRobotHeartbeatPulse := FALSE;

IF GVL_MQTT.bVisuForceDisableTeachIndicator THEN
	bRobotArmTeachMode := FALSE;
END_IF

END_FUNCTION_BLOCK

// ---- POUs/F_ParseStateDisplay.TcPOU
FUNCTION F_ParseStateDisplay : STRING(255)
VAR_INPUT
	{attribute 'TcEncoding':='UTF-8'}
	sPayload		: STRING(255);
END_VAR
VAR
	nStartPos	: INT;
	nEndPos		: INT;
	nPartLen	: INT;
END_VAR

F_ParseStateDisplay := sPayload;

nStartPos := FIND(sPayload, '"state":"');
IF nStartPos > 0 THEN
	nStartPos := nStartPos + 9;
	nEndPos := FIND(sPayload, '","');
	IF nEndPos = 0 THEN
		nEndPos := FIND(sPayload, '"}');
	END_IF

	nPartLen := nEndPos - nStartPos;
	IF nPartLen > 0 THEN
		F_ParseStateDisplay := MID(sPayload, nPartLen, nStartPos);
	END_IF
END_IF

END_FUNCTION

// ---- POUs/F_ParseErrorDisplay.TcPOU
FUNCTION F_ParseErrorDisplay : STRING(255)
VAR_INPUT
	{attribute 'TcEncoding':='UTF-8'}
	sPayload		: STRING(255);
END_VAR
VAR
	nStartPos	: INT;
	nEndPos		: INT;
	nPartLen	: INT;
	sParsed		: STRING(255);
END_VAR

F_ParseErrorDisplay := sPayload;

IF FIND(sPayload, '"error":false') > 0 THEN
	F_ParseErrorDisplay := 'OK';
ELSIF FIND(sPayload, '"error":true') > 0 THEN
	nStartPos := FIND(sPayload, '"message":"');
	IF nStartPos > 0 THEN
		nStartPos := nStartPos + 11;
		nEndPos := FIND(sPayload, '"}');
		nPartLen := nEndPos - nStartPos;
		IF nPartLen > 0 THEN
			sParsed := MID(sPayload, nPartLen, nStartPos);
			IF LEN(sParsed) > 0 THEN
				F_ParseErrorDisplay := sParsed;
			ELSE
				F_ParseErrorDisplay := 'ERROR';
			END_IF
		ELSE
			F_ParseErrorDisplay := 'ERROR';
		END_IF
	ELSE
		F_ParseErrorDisplay := 'ERROR';
	END_IF
END_IF

END_FUNCTION

// ---- POUs/FB_QrVision.TcPOU
FUNCTION_BLOCK FB_QrVision
VAR_INPUT
  bEnable : BOOL := TRUE;
END_VAR
VAR_OUTPUT
  bCodeFound    : BOOL := FALSE;
  sCodeAsString : STRING(255) := '';
  sDisplayText  : STRING(512) := '';
  hrLast        : HRESULT := 0;
  bCameraConnected : BOOL := FALSE;
END_VAR
VAR
  fbCameraControl   : FB_VN_GevCameraControl;
  eState            : ETcVnCameraState;
  hr                : HRESULT;

  ipImageIn         : ITcVnImage;
  ipImageInDisp     : ITcVnDisplayableImage;
  ipImageRGB        : ITcVnImage;
  ipImageResDisp    : ITcVnDisplayableImage;

  ipCodeDecodedList : ITcVnContainer;
  ipCodeContourList : ITcVnContainer;
  hrQr              : HRESULT;
  nQrAttempt        : USINT;

  aColorRed         : TcVnVector4_LREAL := [255, 0, 0, 255];
END_VAR

eState := fbCameraControl.GetState();

// Camera connected when opened or acquiring
IF (eState = TCVN_CS_OPENED) OR (eState = TCVN_CS_STARTACQUISITION) OR (eState = TCVN_CS_ACQUIRING) THEN
  bCameraConnected := TRUE;
ELSE
  bCameraConnected := FALSE;
END_IF

CASE eState OF
  TCVN_CS_ERROR:
    fbCameraControl.Reset();

  TCVN_CS_INITIAL,
  TCVN_CS_OPENING,
  TCVN_CS_OPENED,
  TCVN_CS_STARTACQUISITION:
    IF bEnable THEN
      hr := fbCameraControl.StartAcquisition();
    END_IF

  TCVN_CS_ACQUIRING:
    IF bEnable THEN
      hr := fbCameraControl.GetCurrentImage(ipImageIn);

      IF SUCCEEDED(hr) AND ipImageIn <> 0 THEN
        hr := F_VN_CopyIntoDisplayableImage(ipImageIn, ipImageInDisp, hr);

        bCodeFound := FALSE;
        sCodeAsString := '';
        sDisplayText := '';
        ipCodeDecodedList := 0;
        ipCodeContourList := 0;

        FOR nQrAttempt := 1 TO 3 DO
          hrQr := 0;

          CASE nQrAttempt OF
            1:
              hrQr := F_VN_ReadQRCodeExp(
                ipSrcImage      := ipImageIn,
                ipDecodedData   := ipCodeDecodedList,
                ipContours      := ipCodeContourList,
                nCodeNumber     := 1,
                eSearchStrategy := TCVN_CSS_ONLY_NOT_INVERTED + TCVN_CSS_ONLY_NOT_FLIPPED,
                hrPrev          := hrQr
              );
            2:
              hrQr := F_VN_ReadQRCodeExp(
                ipSrcImage      := ipImageIn,
                ipDecodedData   := ipCodeDecodedList,
                ipContours      := ipCodeContourList,
                nCodeNumber     := 1,
                eSearchStrategy := TCVN_CSS_ONLY_NOT_FLIPPED,
                hrPrev          := hrQr
              );
            3:
              hrQr := F_VN_ReadQRCodeExp(
                ipSrcImage      := ipImageIn,
                ipDecodedData   := ipCodeDecodedList,
                ipContours      := ipCodeContourList,
                nCodeNumber     := 1,
                eSearchStrategy := TCVN_CSS_ONLY_NOT_INVERTED,
                hrPrev          := hrQr
              );
          END_CASE

          IF SUCCEEDED(hrQr) AND ipCodeDecodedList <> 0 THEN
            bCodeFound := TRUE;
            hr := F_VN_ExportSubContainer_String(ipCodeDecodedList, 0, sCodeAsString, 255, hr);
            EXIT;
          END_IF
        END_FOR

        hr := F_VN_ConvertColorSpace(ipImageIn, ipImageRGB, TCVN_CST_GRAY_TO_RGB, hr);

        IF bCodeFound AND ipCodeContourList <> 0 THEN
          hr := F_VN_DrawContours(ipCodeContourList, 0, ipImageRGB, aColorRed, 3, hr);
          sDisplayText := CONCAT('QR: ', sCodeAsString);
        ELSE
          sDisplayText := 'No QR Code Found';
        END_IF

        hr := F_VN_PutTextExp(sDisplayText, ipImageRGB, 50, 100, ETcVnFontType.TCVN_FT_HERSHEY_SIMPLEX, 1.0, aColorRed, 2, TCVN_LT_8_CONNECTED, FALSE, hr);
        hr := F_VN_CopyIntoDisplayableImage(ipImageRGB, ipImageResDisp, hr);
      END_IF
    ELSE
      bCodeFound := FALSE;
      sCodeAsString := '';
        sDisplayText := 'QR scanner OFF';
    END_IF

  TCVN_CS_STOPACQUISITION:
    ;
  TCVN_CS_TRIGGERING:
    ;
  TCVN_CS_CLOSING:
    ;
END_CASE

hrLast := hr;

END_FUNCTION_BLOCK

// ---- GlobalTextList.TcGTLO
TEXTLIST GlobalTextList
  655 = 'Actibe'
  56 = 'Active'
  14 = 'Broker Host'
  493 = 'Broker Host: %s'
  78 = 'Broker Port'
  225 = 'Broker Port: %s'
  229 = 'Broker: %s'
  314 = 'Conncted'
  184 = 'Connected'
  798 = 'Current State : %s'
  156 = 'Current State: %s'
  520 = 'Display: '
  981 = 'Display: %s'
  309 = 'Done'
  631 = 'E-STOP'
  797 = 'EMERGENCY STOP'
  682 = 'Enable Auto'
  297 = 'Enable MQTT'
  906 = 'Enable QR'
  308 = 'Enable QrVision'
  904 = 'Enabled'
  818 = 'Error'
  705 = 'Found'
  9 = 'GOTO '
  576 = 'GOTO Camera'
  299 = 'GOTO Discard'
  667 = 'GOTO Inductieve'
  837 = 'GOTO Mixer'
  584 = 'GOTO Scale'
  207 = 'Heartbeat status'
  443 = 'Heartbeat status: %s'
  523 = 'Inductieve Sensor'
  638 = 'Last Acknowledgement : %s'
  954 = 'Metaal Detectie'
  717 = 'Mixer'
  803 = 'MixerCmd: %s'
  227 = 'MixerCmdRaw: %s'
  736 = 'MixerError: %s'
  519 = 'MixerErrorRaw: %s'
  163 = 'MixerState: %s'
  767 = 'MixerStateRaw: %s'
  369 = 'MQTT Broker'
  28 = 'MQTT Monitor'
  831 = 'Online'
  66 = 'OTO Camera'
  503 = 'QR Code: %s'
  501 = 'QR Enabled: %s'
  494 = 'QR Enabled: %s '
  502 = 'QR Found: %s'
  504 = 'QR Status: %s'
  232 = 'QrVision'
  441 = 'Robot Arm'
  370 = 'RobotCmd: %s'
  200 = 'RobotCmdRaw: %s'
  878 = 'RobotError: %s'
  462 = 'RobotErrorRaw: %s'
  122 = 'RobotState: %s'
  304 = 'RobotStateRaw: %s'
  621 = 'Running'
  390 = 'Save'
  29 = 'SAVE POSITION'
  740 = 'Start'
  619 = 'Start Auto'
  742 = 'Start Robot'
  600 = 'StartKnop'
  916 = 'Startknop'
  632 = 'Status'
  257 = 'Stop'
  377 = 'Stopknop'
  591 = 't'
  992 = 'Teach'
  982 = 'Teach Camera'
  10 = 'Teach Discard'
  480 = 'Teach Inductieve'
  2 = 'Teach Mixer'
  315 = 'TEACH MODE'
  948 = 'Teach Scale'
  865 = 'Transportband'
  930 = 'Vision Done'
END_TEXTLIST

// ---- VISUs/PannenkoekenDashboard.TcVIS
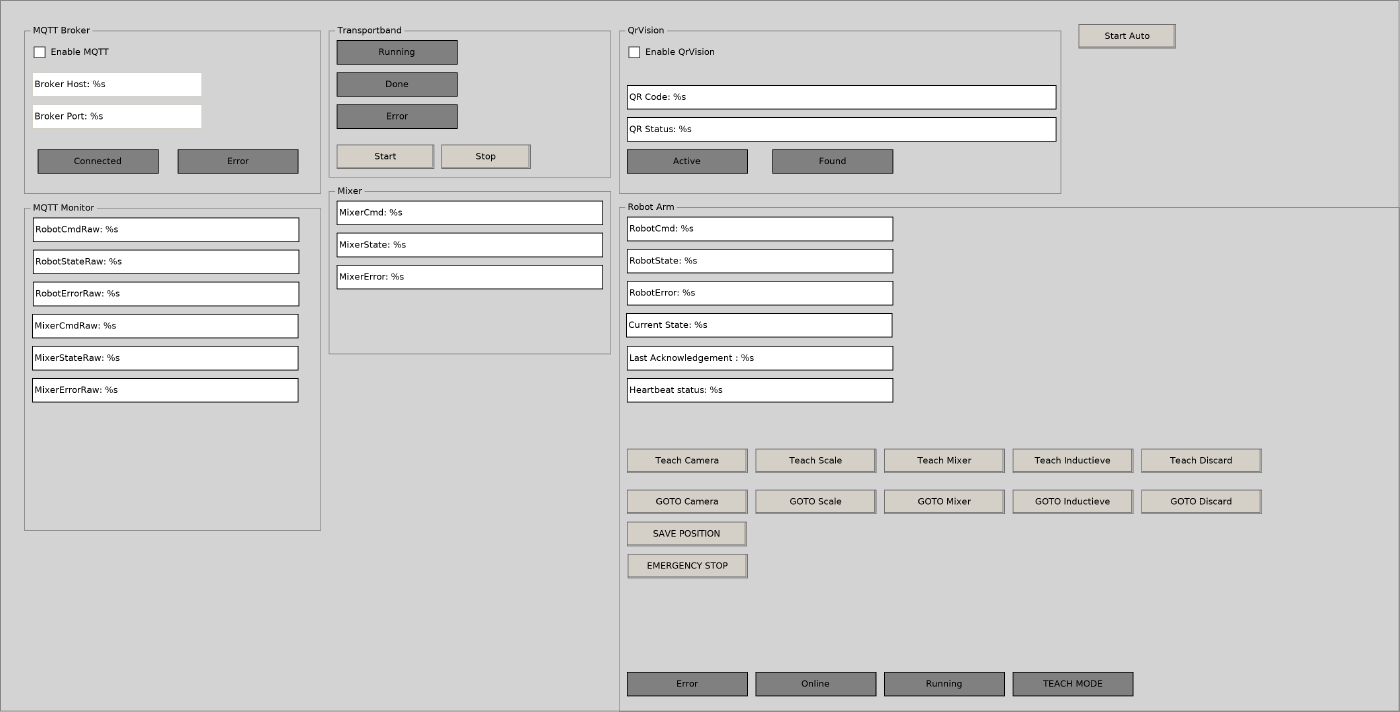
VISUALIZATION PannenkoekenDashboard  // 1742x887
    GroupBox (30,30 369x211), "MQTT Broker"
        Checkbox (10,20 150x30), "Enable MQTT", variable: GVL_MQTT.bEnableMqtt
        Rectangle (191,156 150x30), "Error"
        Rectangle (17,156 150x30), "Connected", colour toggle: GVL_MQTT.bMqttConnected
        Textfield (10,60 211x30), "Broker Host: %s", text variable: GVL_MQTT.sMqttBroker
        Textfield (10,100 211x30), "Broker Port: %s", text variable: GVL_MQTT.nMqttPort
    GroupBox (30,251 369x410), "MQTT Monitor"
        Rectangle (10,140 331x30), "MixerCmdRaw: %s", text variable: GVL_MQTT.sMixerCmdRaw
        Rectangle (10,180 331x30), "MixerStateRaw: %s", text variable: GVL_MQTT.sMixerStateRaw
        Rectangle (10,220 331x30), "MixerErrorRaw: %s", text variable: GVL_MQTT.sMixerErrorRaw
        Rectangle (11,20 331x30), "RobotCmdRaw: %s", text variable: GVL_MQTT.sRobotCmdRaw
        Rectangle (11,60 331x30), "RobotStateRaw: %s", text variable: GVL_MQTT.sRobotStateRaw
        Rectangle (11,100 331x30), "RobotErrorRaw: %s", text variable: GVL_MQTT.sRobotErrorRaw
    GroupBox (770,250 972x637), "Robot Arm"
        Rectangle (10,20 331x30), "RobotCmd: %s", text variable: GVL_MQTT.sRobotCmdDisplay
        Rectangle (10,60 331x30), "RobotState: %s", text variable: GVL_MQTT.sRobotStateDisplay
        Rectangle (10,100 331x30), "RobotError: %s", text variable: GVL_MQTT.sRobotErrorDisplay
        Rectangle (10,587 150x30), "Error", colour toggle: GVL_MQTT.bRobotArmAlarm
        Rectangle (170,587 150x30), "Online", colour toggle: GVL_MQTT.bRobotArmOnline
        Rectangle (330,587 150x30), "Running", colour toggle: GVL_MQTT.bRobotArmBusy
        Rectangle (10,221 331x30), "Heartbeat status: %s", text variable: GVL_MQTT.sRobotHeartbeatDisplay
        Rectangle (9,140 331x30), "Current State: %s", text variable: GVL_MQTT.sRobotArmDisplay
        Button (10,309 150x30), "Teach Camera"
            OnMouseClick: execute { GVL_MQTT.sRobotTargetPose := 'camera'; GVL_MQTT.bVisuRobotTeach  := TRUE; }
        Button (170,309 150x30), "Teach Scale"
            OnMouseClick: execute { GVL_MQTT.sRobotTargetPose := 'scale'; GVL_MQTT.bVisuRobotTeach  := TRUE; }
        Button (330,309 150x30), "Teach Mixer"
            OnMouseClick: execute { GVL_MQTT.sRobotTargetPose := 'mixer'; GVL_MQTT.bVisuRobotTeach  := TRUE; }
        Button (490,309 150x30), "Teach Inductieve"
            OnMouseClick: execute { GVL_MQTT.sRobotTargetPose := 'inductive'; GVL_MQTT.bVisuRobotTeach  := TRUE; }
        Button (650,309 150x30), "Teach Discard"
            OnMouseClick: execute { GVL_MQTT.sRobotTargetPose := 'discard'; GVL_MQTT.bVisuRobotTeach  := TRUE; }
        Button (10,360 150x30), "GOTO Camera"
            OnMouseClick: execute { GVL_MQTT.sRobotTargetPose := 'camera'; GVL_MQTT.bVisuRobotGoto   := TRUE; }
        Button (10,400 149x30), "SAVE POSITION"
            tap GVL_MQTT.bVisuRobotSave
        Button (11,440 149x30), "EMERGENCY STOP"
            tap GVL_MQTT.bVisuRobotStop
        Rectangle (10,181 331x30), "Last Acknowledgement : %s", text variable: GVL_MQTT.sRobotArmAck
        Rectangle (490,587 150x30), "TEACH MODE", colour toggle: GVL_MQTT.bRobotArmTeachMode
    GroupBox (409,30 351x191), "Transportband"
        Button (10,150 121x30), "Start"
            tap GVL_MQTT.bVisuStartTransportband
        Button (140,150 111x30), "Stop"
            tap GVL_MQTT.bVisuStopTransportband
        Rectangle (10,20 150x30), "Running", colour toggle: GVL_MQTT.bTransportbandRunning
        Rectangle (10,60 150x30), "Done", colour toggle: GVL_MQTT.bTransportbandDone
        Rectangle (10,100 150x30), "Error", colour toggle: GVL_MQTT.bSystemError
    GroupBox (409,230 351x211), "Mixer"
        Rectangle (10,60 331x30), "MixerState: %s", text variable: GVL_MQTT.sMixerStateDisplay
        Rectangle (10,20 331x30), "MixerCmd: %s", text variable: GVL_MQTT.sMixerCmdDisplay
        Rectangle (10,100 331x30), "MixerError: %s", text variable: GVL_MQTT.sMixerErrorDisplay
    GroupBox (770,30 550x211), "QrVision"
        Rectangle (10,76 534x30), "QR Code: %s", text variable: GVL_Data.sQrCodeText
        Rectangle (10,116 534x30), "QR Status: %s", text variable: GVL_Data.sQrDisplayText
        Rectangle (10,156 150x30), "Active", colour toggle: GVL_Data.bQrActive
        Rectangle (191,156 150x30), "Found", colour toggle: GVL_Data.bQrCodeFound
        Checkbox (10,20 150x30), "Enable QrVision", variable: GVL_Data.bQrEnabled
    Button (940,610 150x30), "GOTO Scale"
        OnMouseClick: execute { GVL_MQTT.sRobotTargetPose := 'scale'; GVL_MQTT.bVisuRobotGoto   := TRUE; }
    Button (1100,610 150x30), "GOTO Mixer"
        OnMouseClick: execute { GVL_MQTT.sRobotTargetPose := 'mixer'; GVL_MQTT.bVisuRobotGoto   := TRUE; }
    Button (1260,610 150x30), "GOTO Inductieve"
        OnMouseClick: execute { GVL_MQTT.sRobotTargetPose := 'inductive'; GVL_MQTT.bVisuRobotGoto   := TRUE; }
    Button (1420,610 150x30), "GOTO Discard"
        OnMouseClick: execute { GVL_MQTT.sRobotTargetPose := 'discard'; GVL_MQTT.bVisuRobotGoto   := TRUE; }
    Button (1342,30 121x30), "Start Auto"
        tap GVL_MQTT.bVisuStartSequence
END_VISUALIZATION
